(* IEC 61131-3 sources: llm-plc-st-eval/codesys/dobles/B7, 9 files *)

(* ---- 01_Correcta.st ---- *)
(* DOBLE DE PRUEBA B7/Correcta - NO ES CORPUS. Esperado: veredicto 1 *)
FUNCTION SelBomba : BOOL
VAR_INPUT
    modoAuto : BOOL;
    btnManual : BOOL;
    nivelBajo : BOOL;
END_VAR
IF modoAuto THEN
    SelBomba := nivelBajo;
ELSE
    SelBomba := btnManual;
END_IF
END_FUNCTION

(* ---- 04_ModoInvertido.st ---- *)
(* DOBLE DE PRUEBA B7/ModoInvertido - NO ES CORPUS. Esperado: veredicto 2, falla en el paso 1 *)
FUNCTION SelBomba : BOOL
VAR_INPUT
    modoAuto : BOOL;
    btnManual : BOOL;
    nivelBajo : BOOL;
END_VAR
IF modoAuto THEN
    SelBomba := btnManual;
ELSE
    SelBomba := nivelBajo;
END_IF
END_FUNCTION

(* ---- 05_OrSimple.st ---- *)
(* DOBLE DE PRUEBA B7/OrSimple - NO ES CORPUS. Esperado: veredicto 2, falla en el paso 3 *)
FUNCTION SelBomba : BOOL
VAR_INPUT
    modoAuto : BOOL;
    btnManual : BOOL;
    nivelBajo : BOOL;
END_VAR
SelBomba := btnManual OR nivelBajo;
END_FUNCTION

(* ---- 06_NivelInvertido.st ---- *)
(* DOBLE DE PRUEBA B7/NivelInvertido - NO ES CORPUS. Esperado: veredicto 2, falla en el paso 4 *)
FUNCTION SelBomba : BOOL
VAR_INPUT
    modoAuto : BOOL;
    btnManual : BOOL;
    nivelBajo : BOOL;
END_VAR
IF modoAuto THEN
    SelBomba := NOT nivelBajo;
ELSE
    SelBomba := btnManual;
END_IF
END_FUNCTION

(* ---- 07_BotonTambienEnAuto.st ---- *)
(* DOBLE DE PRUEBA B7/BotonTambienEnAuto - NO ES CORPUS. Esperado: veredicto 2, falla en el paso 6 *)
FUNCTION SelBomba : BOOL
VAR_INPUT
    modoAuto : BOOL;
    btnManual : BOOL;
    nivelBajo : BOOL;
END_VAR
IF modoAuto THEN
    SelBomba := nivelBajo OR btnManual;
ELSE
    SelBomba := btnManual;
END_IF
END_FUNCTION

(* ---- 02_CorrectaFB.st ---- *)
(* DOBLE DE PRUEBA B7/CorrectaFB - NO ES CORPUS. Esperado: veredicto 1 *)
FUNCTION_BLOCK SelBomba
VAR_INPUT
    modoAuto : BOOL;
    btnManual : BOOL;
    nivelBajo : BOOL;
END_VAR
VAR_OUTPUT
    bomba : BOOL;
END_VAR
VAR
    nada : BOOL;
END_VAR
IF modoAuto THEN
    bomba := nivelBajo;
ELSE
    bomba := btnManual;
END_IF
END_FUNCTION_BLOCK

(* ---- 08_MemoriaEnAuto.st ---- *)
(* DOBLE DE PRUEBA B7/MemoriaEnAuto - NO ES CORPUS. Esperado: veredicto 2, falla en el paso 5 *)
FUNCTION_BLOCK SelBomba
VAR_INPUT
    modoAuto : BOOL;
    btnManual : BOOL;
    nivelBajo : BOOL;
END_VAR
VAR_OUTPUT
    bomba : BOOL;
END_VAR
VAR
    nada : BOOL;
END_VAR
IF modoAuto THEN
    bomba := bomba OR nivelBajo;
ELSE
    bomba := btnManual;
END_IF
END_FUNCTION_BLOCK

(* ---- 03_CorrectaPRG.st ---- *)
(* DOBLE DE PRUEBA B7/CorrectaPRG - NO ES CORPUS. Esperado: veredicto 1 *)
PROGRAM SelBomba
VAR_INPUT
    modoAuto : BOOL;
    btnManual : BOOL;
    nivelBajo : BOOL;
END_VAR
VAR_OUTPUT
    bomba : BOOL;
END_VAR
VAR
    nada : BOOL;
END_VAR
IF modoAuto THEN
    bomba := nivelBajo;
ELSE
    bomba := btnManual;
END_IF
END_PROGRAM

(* ---- 09_TelerruptorManual.st ---- *)
(* DOBLE DE PRUEBA B7/TelerruptorManual - NO ES CORPUS. Esperado: veredicto 2, falla en el paso 2 *)
PROGRAM SelBomba
VAR_INPUT
    modoAuto : BOOL;
    btnManual : BOOL;
    nivelBajo : BOOL;
END_VAR
VAR_OUTPUT
    bomba : BOOL;
END_VAR
VAR
    prev : BOOL;
END_VAR
IF modoAuto THEN
    bomba := nivelBajo;
ELSIF btnManual AND NOT prev THEN
    bomba := NOT bomba;
END_IF
prev := btnManual;
END_PROGRAM
